// TIA Portal V20 export
// export: Created 2026-10-19T18:42:07.4796645Z, ExportSetting WithDefaults, DisplayName Totally Integrated Automation Portal, DisplayVersion V20 Update 6, DisplayName TIA Portal Openness, DisplayVersion V20 Update 6, DisplayName TIA Portal Version Control Interface, DisplayVersion V20 Update 6, DisplayName SINAMICS Startdrive Advanced, DisplayVersion V20 SP1, DisplayName SINAMICS Startdrive G130, G150, S120, S150, SINAMICS MV, G220, S200, S210, DisplayVersion V20 SP1, DisplayName SINAMICS Startdrive G110M, G120, G120C, G120D, G120P, G115D, DisplayVersion V20 SP1, DisplayName STEP 7 Professional, DisplayVersion V20 Update 6, DisplayName STEP 7 Safety, DisplayVersion V20 Update 2, DisplayName WinCC Basic/Comfort/Advanced, DisplayVersion V20 Update 6, DisplayName WinCC Unified, DisplayVersion V20 Update 6
DATA_BLOCK "Watchdog_Settings"   // DB134
{ S7_Optimized_Access := 'TRUE' }
VERSION : 0.1
// stored: AutoNumber true, DBAccessibleFromOPCUA true, InstanceOfName Watchdog_Settings_UDT, InstanceOfType UDT, IsOnlyStoredInLoadMemory false, IsWriteProtectedInAS false
"Watchdog_Settings_UDT"
   // VAR
   //    VTD : UDInt := 500;
   //    EConveyor : UDInt := 500;
   //    Cnv2_Buffer_L : Array[2..5] of UDInt;
   //    Cnv1_Buffer_L : Array[2..5] of UDInt;
   //    Pallet_INOut : UDInt := 500;
   //    Shuttle_INOut : UDInt := 500;
   //    Level_2 : UDInt;
   //    Level_3 : UDInt;
   //    Level_4 : UDInt;
   //    Level_5 : UDInt;
   //    Level_6 : UDInt;
   // END_VAR
BEGIN
END_DATA_BLOCK
